FUNCTION_BLOCK ThermometerS (* Composite Function Block Type *)
  (* Standard: 61499-2 *)
  (* Version 0.0, 6/21/2016, Andrei, nxtControl GmbH, template *)
  PACKAGE Main;
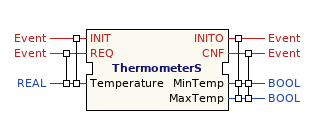
  EVENT_INPUT
    INIT WITH Temperature; (* Initialization Request *)
    REQ WITH Temperature; (* Normal Execution Request *)
  END_EVENT
  EVENT_OUTPUT
    INITO WITH MinTemp, MaxTemp; (* Initialization Confirm *)
    CNF WITH MinTemp, MaxTemp; (* Execution Confirmation *)
  END_EVENT
  VAR_INPUT
    Temperature : REAL; (* Input event qualifier *)
  END_VAR
  VAR_OUTPUT
    MinTemp : BOOL; (* Output event qualifier *)
    MaxTemp : BOOL;
  END_VAR
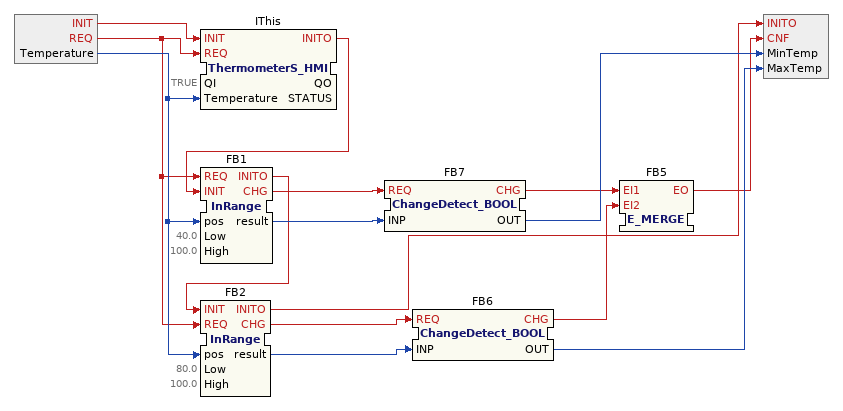
  FBS
    IThis : ThermometerS_HMI(QI := TRUE);
    FB1 : InRange(Low := 40.0, High := 100.0);
    FB2 : InRange(Low := 80.0, High := 100.0);
    FB5 : E_MERGE;
    FB6 : ChangeDetect_BOOL;
    FB7 : ChangeDetect_BOOL;
  END_FBS
  EVENT_CONNECTIONS
    INIT TO IThis.INIT;
    REQ TO IThis.REQ;
    REQ TO FB1.REQ;
    IThis.INITO TO FB1.INIT;
    FB1.INITO TO FB2.INIT;
    FB2.INITO TO INITO;
    FB2.CHG TO FB6.REQ;
    FB1.CHG TO FB7.REQ;
    FB7.CHG TO FB5.EI1;
    FB6.CHG TO FB5.EI2;
    FB5.EO TO CNF;
    REQ TO FB2.REQ;
  END_CONNECTIONS
  DATA_CONNECTIONS
    Temperature TO FB1.pos;
    Temperature TO FB2.pos;
    Temperature TO IThis.Temperature;
    FB2.result TO FB6.INP;
    FB6.OUT TO MaxTemp;
    FB1.result TO FB7.INP;
    FB7.OUT TO MinTemp;
  END_CONNECTIONS
END_FUNCTION_BLOCK
